// TIA Portal V21 export
// export: Created 2026-11-11T00:48:23.1848694Z, ExportSetting WithDefaults, DisplayName Totally Integrated Automation Portal, DisplayVersion V21 Update 3, DisplayName STEP 7 Professional, DisplayVersion V21 Update 3, DisplayName STEP 7 Safety, DisplayVersion V21, DisplayName Tech WebApplication, DisplayVersion V21, DisplayName WinCC Basic/Comfort/Advanced, DisplayVersion V21 Update 3, DisplayName WinCC Unified, DisplayVersion V21 Update 3
FUNCTION_BLOCK "FB_Scl_sl112"   // FB196, SCL
{ S7_Optimized_Access := 'TRUE' }
VERSION : 0.1
// stored: AutoNumber true, IsIECCheckEnabled false, IsRetainMemResEnabled false, MemoryReserve 100, SetENOAutomatically false, UDAEnableTagReadback false
   VAR_INPUT
      v_reset : Bool;
      v_jog : Bool;
      v_drum_en : Bool;
      v_lst_step : Byte;
   END_VAR
   VAR_OUTPUT
      v_q : Bool;
      v_out_word : Word;
      v_err_code : Word;
   END_VAR
   VAR
      inst { S7_SetPoint := 'True'} : DRUM;
   END_VAR
BEGIN
   #inst(RESET := #v_reset, JOG := #v_jog, DRUM_EN := #v_drum_en, LST_STEP := #v_lst_step, Q => #v_q, OUT_WORD => #v_out_word, ERR_CODE => #v_err_code);
END_FUNCTION_BLOCK
